// TIA Portal V21 export
// export: Created 2000-01-01T00:00:00.0000000Z, ExportSetting None
TYPE "UDT_HMI_AnalogScale"
   STRUCT
      bManualOverride { ExternalWritable := 'False'} : Bool;   // HMI手动仿真覆盖使能
      bResetCmd { ExternalWritable := 'False'} : Bool;   // HMI故障与锁存报警复位触发
      rManualValue { ExternalWritable := 'False'} : Real;   // HMI手动强制工程值给定
      rRawMin { ExternalWritable := 'False'} : Real;   // 原始码值下限（默认 0.0 或 5530.0）
      rRawMax { ExternalWritable := 'False'} : Real;   // 原始码值上限（默认 27648.0）
      rEngMin { ExternalWritable := 'False'} : Real;   // 工程量下限（如 0.0）
      rEngMax { ExternalWritable := 'False'} : Real;   // 工程量上限（如 100.0）
      rLimitHH { ExternalWritable := 'False'} : Real;   // 高高限报警阈值
      rLimitH { ExternalWritable := 'False'} : Real;   // 高限警告阈值
      rLimitL { ExternalWritable := 'False'} : Real;   // 低限警告阈值
      rLimitLL { ExternalWritable := 'False'} : Real;   // 低低限报警阈值
      rScaledValue { ExternalWritable := 'False'} : Real;   // 状态反馈：当前标定工程值
      bAlarmHH { ExternalWritable := 'False'} : Bool;   // 状态反馈：高高限报警
      bAlarmH { ExternalWritable := 'False'} : Bool;   // 状态反馈：高限报警
      bAlarmL { ExternalWritable := 'False'} : Bool;   // 状态反馈：低限报警
      bAlarmLL { ExternalWritable := 'False'} : Bool;   // 状态反馈：低低限报警
      bWireBreak { ExternalWritable := 'False'} : Bool;   // 状态反馈：断线或溢出故障
      wStatus { ExternalWritable := 'False'} : Word;   // 故障码：16#0000正常, 16#8200量程除零, 16#8201阈值顺序错, 16#8401断线/溢出
   END_STRUCT;
END_TYPE
